# EPICS substitutions: niusb/niusbApp/Db/USB6210.substitutions
# The USB-6210: every record, by measComp's names. Macros: P, PORT, MAX_POINTS (from the entity); the templates at the image's /epics/support/niusb/db.
file "/epics/support/niusb/db/niusbDevice.template" { pattern {} {} }

file "/epics/support/niusb/db/niusbAi.template"
{
pattern
{ N, ADDR }
{ 1, 0 }
{ 2, 1 }
{ 3, 2 }
{ 4, 3 }
{ 5, 4 }
{ 6, 5 }
{ 7, 6 }
{ 8, 7 }
{ 9, 8 }
{ 10, 9 }
{ 11, 10 }
{ 12, 11 }
{ 13, 12 }
{ 14, 13 }
{ 15, 14 }
{ 16, 15 }
}

file "/epics/support/niusb/db/niusbBi.template"
{
pattern
{ N, LINE, MASK }
{ 1, 0, 0x1 }
{ 2, 1, 0x2 }
{ 3, 2, 0x4 }
{ 4, 3, 0x8 }
}

file "/epics/support/niusb/db/niusbBo.template"
{
pattern
{ N, LINE, MASK }
{ 1, 0, 0x1 }
{ 2, 1, 0x2 }
{ 3, 2, 0x4 }
{ 4, 3, 0x8 }
}

file "/epics/support/niusb/db/niusbWaveDig.template" { pattern {} {} }

file "/epics/support/niusb/db/niusbWaveDigN.template"
{
pattern
{ N, ADDR }
{ 1, 0 }
{ 2, 1 }
{ 3, 2 }
{ 4, 3 }
{ 5, 4 }
{ 6, 5 }
{ 7, 6 }
{ 8, 7 }
{ 9, 8 }
{ 10, 9 }
{ 11, 10 }
{ 12, 11 }
{ 13, 12 }
{ 14, 13 }
{ 15, 14 }
{ 16, 15 }
}
